TYPE ST_VFD_DRIVE_REF : FB_VFD_Drive_REF;
END_TYPE

(* stored: Version 1.1.0.1, ProductVersion 3.1.4024.15
   DUT ST_VFD_DRIVE_REF: Id {8533ef6a-a345-411e-b925-c14ab17ffe90} *)
